Fanuc KAREL source: KO00017.KL

PROGRAM KO00017
%NOLOCKGROUP
VAR
  P1: XYZWPREXT
  P2: XYZWPREXT
  P3: XYZWPREXT
  OUT: POSITION
BEGIN
  OUT = FRAME(P1, P2, P3)
END KO00017
